FUNCTION FC_TransformPosition : LREAL
VAR_INPUT
	fOffset: LREAL;
	fPosition: LREAL;
END_VAR

FC_TransformPosition:=fOffset+fPosition;

END_FUNCTION

(* stored: Version 1.1.0.1, ProductVersion 3.1.4024.12
   POU FC_TransformPosition: Id {458779fb-96d1-4daa-8f50-1fb794fac52b}, SpecialFunc None *)
